Fanuc KAREL source: KA00102.KL

PROGRAM KA00102
%NOLOCKGROUP
VAR
  SRC: VECTOR
  DST: XYZWPR
BEGIN
  SRC.X = 1.0
  DST = SRC
END KA00102
